// TIA Portal V21 export
DATA_BLOCK "Signalläuchte_DB"   // DB13
// stored: InstanceOfName Signalläuchte, InstanceOfType FB
"Signalläuchte"
   // VAR
   //    blink_start : Bool;
   //    state : Int;
   // END_VAR
BEGIN
END_DATA_BLOCK
